// TIA Portal V20 export
// export: Created 2026-10-12T04:58:21.5153537Z, ExportSetting WithDefaults, DisplayName Totally Integrated Automation Portal, DisplayVersion V20, DisplayName TIA Portal Openness, DisplayVersion V20, DisplayName TIA Portal Teamcenter Gateway, DisplayVersion V20, DisplayName TIA Portal Version Control Interface, DisplayVersion V20, DisplayName SINAMICS Startdrive Advanced, DisplayVersion V20 SP1 Update 2, DisplayName SINAMICS Startdrive G110M, G120, G120C, G120D, G120P, G115D, DisplayVersion V20 SP1 Update 2, DisplayName SINAMICS Startdrive G130, G150, S120, S150, SINAMICS MV, G220, S200, S210, DisplayVersion V20 SP1 Update 2, DisplayName STEP 7 Professional, DisplayVersion V20, DisplayName STEP 7 Safety, DisplayVersion V20, DisplayName WinCC Basic/Comfort/Advanced, DisplayVersion V20, DisplayName WinCC Professional, DisplayVersion V20, DisplayName WinCC Unified, DisplayVersion V20
FUNCTION "FRK_ConfigBoot" : Void   // FC103, SCL
{ S7_Optimized_Access := 'TRUE' }
VERSION : 0.1
// stored: AutoNumber true, IsIECCheckEnabled false, SetENOAutomatically false, UDAEnableTagReadback false
   VAR_INPUT
      Startup : Bool;
   END_VAR
   VAR_TEMP
      Index : Int;
   END_VAR
BEGIN

   IF NOT #Startup THEN
       RETURN;
   END_IF;
   "FRK_ConfigRuntime".Fresh := "FRK_ConfigStore".SchemaVersion = 0;
   IF "FRK_ConfigStore".SchemaVersion <> 1 THEN
       FOR #Index := 1 TO 114 DO
           "FRK_ConfigStore".Rows[#Index].Used := FALSE;
       END_FOR;
       IF NOT "FRK_ConfigRuntime".Fresh THEN
           "FRK_ConfigLoss"(RootIndex := 1,
                            Scope := 'StationA');
       END_IF;
       "FRK_ConfigStore".ActiveModels[1] := 'MODEL_A';
       IF NOT "FRK_ConfigRuntime".Fresh THEN
           "FRK_ConfigLoss"(RootIndex := 2,
                            Scope := 'StationB');
       END_IF;
       "FRK_ConfigStore".ActiveModels[2] := 'MODEL_A';
       "FRK_ConfigStore".SchemaVersion := 1;
   END_IF;
   IF "FRK_ConfigStore".ActiveModels[1] <> 'MODEL_A' AND "FRK_ConfigStore".ActiveModels[1] <> 'MODEL_B' THEN
       "FRK_ConfigStore".ActiveModels[1] := 'MODEL_A';
       "FRK_ConfigLoss"(RootIndex := 1,
                        Scope := 'StationA');
   END_IF;
   IF "FRK_ConfigStore".ActiveModels[2] <> 'MODEL_A' AND "FRK_ConfigStore".ActiveModels[2] <> 'MODEL_B' THEN
       "FRK_ConfigStore".ActiveModels[2] := 'MODEL_A';
       "FRK_ConfigLoss"(RootIndex := 2,
                        Scope := 'StationB');
   END_IF;
END_FUNCTION
